(* IEC 61131-3 sources: Elmo_Master/Lasal_PRG/Welcon8Axis_EtherCAT_Test_With_RobotAxis/Network/Axis2, 1 file *)

(* ---- ONE_Axis2_Table.st ---- *)
#define OBJECTS_CONFIG

//Define part of class _LMCAxisBase
//#define _DEBUG_MODUS_MUTEX_OFF
//#define _DEBUG_MODUS_ISSYNCHRON
//#define _DEBUG_MODUS_CHECKSWLIMIT
//#define _DEBUG_MODUS_BRAKING

#define _LMCAXIS_NORMOVERRIDE         1000    // Dieser Override-Wert entspricht 100%.
#define _LMCAXIS_MAXOVERRIDE	        1000		// Maximalwert für Override im LMCAXISBASE (kann mit SetParameter verändert werden.)
#define _LMCAXIS_MINOVERRIDE	           0		// Minimalwert für Override im _LMCAxisBase --> damit man mit Minuswerten nicht in die falsche Richtung fahren kann

#define _LMCAXIS_MIN_POS       -16#07000000    // default MINPOS when INITvalue=0
#define _LMCAXIS_MAX_POS        16#07000000    // default MAXPOS when INITvalue=0

#define _LMCAXIS_OVERVFLOW_POS  16#06000000    // MAX POSITION for checking overflow

#define _LMCAXIS_INVALID_POS    16#3FFFFFFF    // Invalid position for calculating the velocity

#define _LMCAXIS_INTERVAL            10            // original = 10

#define _LMCAXIS_MAX_MASTERDELAY     7    // maximum cycles for delaying the coupling to the master

#define _LMCAXIS_RESO_CALBREMS 100

#ifndef _VOID_POS
  #define  _VOID_POS 16#7FFFFFFF
#endif

/////////////////////
// Polynom 5ten Grades
#define _LMCAXIS_Poly_Pos_A     2.5
#define _LMCAXIS_Poly_Pos_B     3.0
#define _LMCAXIS_Poly_Pos_C     1.0

#define LMC_POLYNOM_V0          0                     // CoupleGearPolynom wenn Slave steht
#define LMC_POLYNOM_V           1                     // CoupleGearPolynom wenn Slave fährt

//////////////////////
// Bewegungsrichtungen
#define _LMCAXIS_MOVE_ANY_WAY              0       // beide Richtungen
#define _LMCAXIS_MOVE_NEG_DIR              1       // nur negative Bewegungsrichtung
#define _LMCAXIS_MOVE_SHORTEST_WAY         2       // kürzester Weg (beide Richtungen)
#define _LMCAXIS_MOVE_POS_DIR              3       // nur positive Bewegungsrichtung

//////////////////////
// Mutex
#define MUTEX_NAME_MAX_LENGTH_LMCAXIS     32   //maximale Anzahl an Zeichen für den Mutexnamen
#define MUTEX_NAME_END_LENGTH_LMCAXIS      3
#define STR_MUTEX_NAME_SEPERATOR_LMCAXIS ".."

#define _LMCAXIS_WAITTIMEPOWERON           90sec    // Wartezeit bei PowerOn bis TimeOut entsteht (maximale Kommutierungszeitdauer beim DiasDrive für Linearmotoren sind 86sec)
#define _LMCAXIS_WAITTIMEPOWEROFF           1sec    // Wartezeit bei PowerOff bis TimeOut entsteht

#define _LMCAXIS_Max_V_FILTER_SIZE   100

//////////////////////
// ruckbegrenzter Modus _JERK_PROFILE
#define MIN_SHRINK_FACTOR_4_CORRECTTOEXACTPOS 0.9
#define MAX_SHRINK_FACTOR_4_CORRECTTOEXACTPOS_FAR 1.2
#define MAX_SHRINK_FACTOR_4_CORRECTTOEXACTPOS_NEAR 5.0
#define MAX_SHRINK_FACTOR_4_CORRECTTOEXACTPOS_WINDOW 5.0

#define MAX_TIME_TO_WAIT_4_BRAKING 3.0 //in Ticks
#define MAX_DURATION_WITH_MAX_ACCEL_TO_MASTER 20000  //in Ticks
#define ALLOWED_AJMP_FACTOR 1.1
#define FACTOR_4_ALLOWED_MASTER_ACCEL_PROFILE_COUPLING 1.2
#define ACCEL_FACTOR_4_PROFILE_COUPLING 1.1
#define JERK_FACTOR_4_PROFILE_COUPLING 1.2

//////////////////////
// LREAL Modi
// #define DEBUG_TRAP_DELTA_ACCEL
#define _LMCAXIS_LREAL_EPSILON 0.000001

#ifndef _DINT_MIN
#define _DINT_MIN -2147483648
#endif

#ifndef _DINT_MAX
#define _DINT_MAX 2147483647
#endif

#define _LMCAXIS_MIN_VEL_MOVECMD 1 // minimale programmierbare Geschwindigkeit fuer LREAL-MoveTypes [internal units / sec]

#define _LMCAXIS_SAFEREFERENCE_TIMEOUT          10 SEC
#define _LMCAXIS_SBTACTIVE_TIMEOUT              16 SEC
#define _LMCAXIS_SAFETYASYNCREQUEST_REPEATTIME  200 MS

#define _LMCAXIS_SBT_SAFESTATE_TESTIDLE    16#0
#define _LMCAXIS_SBT_SAFESTATE_TESTDONE    16#6
#define _LMCAXIS_SBT_SAFESTATE_ERROR      16#E0
#define _LMCAXIS_SBT_FUNCSTATE_FINISH        13

#define _LMCAXIS_LMCPROF_NEWINST_STOPMOVE    77

//+++ einbau HP 13.9.2011 +++++++++++++++++++++++++++++++++++++++++++++++++++++++

//////////////////////
// CoupleGearPolynom
#define _LMCAXIS_FACTOR_JMAX         10
#define _LMCAXIS_FACTOR_T_VAL_X      0.80
#define _LMCAXIS_FACTOR_T_VAL_Z      0.80
#define _LMCAXIS_MIN_TICKS           0

//#define REPORT_TRAPEZOIDSPLINE_DISABLED
#undef REPORT_TRAPEZOIDSPLINE_DISABLED

// Formeltest und Test auf numerische Genauigkeit
//#define CHECK_PRECISION

#define PRAEFIX_KILO          (1000.0)
#ifndef CONVERT_SEC_TO_MSEC
  #define CONVERT_SEC_TO_MSEC   (1000.0)
#endif
//+++++++++++++++++++++++++++++++++++++++++++++++++++++++ einbau HP 13.9.2011 +++

#ifndef LMCMODULEBASE_MAX_LOGININDEX
  #define LMCMODULEBASE_MAX_LOGININDEX      9
#endif

// ===================================================================
// defines linked to safety features
// defines from header file DriveSafetyIF.h from HW lib to reduce dependencies

// VERIFY CMDRSP
// General
#define _LMCAXIS_SAFETY_VERCMD_OK                     0x40000000  // Command successfully processed
#define _LMCAXIS_SAFETY_VERCMD_BUSY                   0x0000000B  // Response to command has not yet been recived
#define _LMCAXIS_SAFETY_VERCMD_EXECUTING              0x4000000B  // Commmand ist still beeing processed ins safety FW
#define _LMCAXIS_SAFETY_VERCMD_WRONG_RUNSTATE         0x40000003  // Command not allowed in current state
#define _LMCAXIS_SAFETY_VERCMD_NOT_NEEDED             0x40000004  // Command executed, although no verification is necessary

#define _LMCAXIS_SAFETY_VERCMD_ERROR_ENC_ID_PROG      0x40000005  // Programming of the encoder index failed

#define _LMCAXIS_SAFETY_VERCMD_INCOMPLETE             0x40000001  // Not all axes requiring verification, have been verified
#define _LMCAXIS_SAFETY_VERCMD_ERROR                  0x40000002  // Saving the HDSL verification status has failed

// VERIFY STATE
#define _LMCAXIS_SAFETY_VERSTATE_UNKOWN               0x00000000  // State has not yet been read
#define _LMCAXIS_SAFETY_VERSTATE_BUSY                 0x0000000B  // State is beeing read

#define _LMCAXIS_SAFETY_VERSTATE_NOT_VERIFIED         0x1A8C5E7B  // Axis not verified, verification necessary
#define _LMCAXIS_SAFETY_VERSTATE_SYSTEM_VERIFIED      0x2B9D6F8C  // Entire drive fully verified
#define _LMCAXIS_SAFETY_VERSTATE_NOT_USED             0x30000000  // no verification necessary for this axis, as not configured as Hiperface DSL

#define _LMCAXIS_SAFETY_VERSTATE_VERIFICATION_PENDING 0x30000001  // Verification has been started for this axis, Programming of the encoder index in progress
#define _LMCAXIS_SAFETY_VERSTATE_AXIS_VERIFIED        0x30000002  // Encoder index has been successfully programmed, Verification completed for this axis (Overall verification necessary at the end)

// REFERENCE CMDRSP
// General
#define _LMCAXIS_SAFETY_REFCMD_OK                     0x40000000  // Command successfully processed
#define _LMCAXIS_SAFETY_REFCMD_BUSY                   0x0000000B  // Response to command has not yet been recived
#define _LMCAXIS_SAFETY_REFCMD_PROGRAMMING_FAILED     0x40000002  // The saving of the offset or the referencing status has failed.
#define _LMCAXIS_SAFETY_REFCMD_WRONG_RUNSTATE         0x40000003  // Command not allowed in current state
#define _LMCAXIS_SAFETY_REFCMD_NOT_NEEDED             0x40000004  // Command executed, although no reference is necessary

// For _LMCAXIS_SAFETY__REFCMD_ACKZERO_POS
#define _LMCAXIS_SAFETY_REFCMD_NOT_ALLOWED            0x40000010  // Absolute position referencing was not started, command not yet allowed
#define _LMCAXIS_SAFETY_REFCMD_NO_MOVEMENT            0x40000011  // Position has not moved far enough from the zero position since the start of referencing
#define _LMCAXIS_SAFETY_REFCMD_WRONG_POSITION         0x40000012  // Newly approached zero position deviates more than permitted from initially approached zero position

// REFERENCE STATE
#define _LMCAXIS_SAFETY_REFSTATE_UNKOWN               0x00000000  //

#define _LMCAXIS_SAFETY_REFSTATE_BUSY                 0x0000000B  // State is beeing read

#define _LMCAXIS_SAFETY_STATE_NOT_REFERENCED          0x1A8C5E7B  // Axis not referenced, referencing necessary
#define _LMCAXIS_SAFETY_STATE_AXIS_REFERENCED         0x2B9D6F8C  // Axis fully referenced
#define _LMCAXIS_SAFETY_STATE_NOT_NEEDED              0x30000000  // No referencing necessary for this axis

#define _LMCAXIS_SAFETY_STATE_WAIT_MOVEMENT           0x30000001  // Referencing has been started, it is waiting for the waiting for the current position to move away from the zero position
#define _LMCAXIS_SAFETY_STATE_ACK_PENDING             0x30000002  // Current position far enough away from zero position, it waits for the zero position to be approached again and confirmed
#define _LMCAXIS_SAFETY_STATE_REFERENCE_DONE          0x30000003  // Zero position successfully confirmed, referencing completed

// DRIVE SAFETY PARA STATES
#define _LMCAXIS_SAFETY_UPDATEPARACLASS_STATE                 16#857E
#define _LMCAXIS_SAFETY_UPDATEPARACLASS_STATE_VER_1           1                   //version 1
#define _LMCAXIS_SAFETY_UPDATEPARACLASS_STATE_VER_MAX         _LMCAXIS_SAFETY_UPDATEPARACLASS_STATE_VER_1   //newest implemented version

#define _LMCAXIS_SAFETY_UPDATEPARACLASS_STATE_GENERAL_ERROR                 1
#define _LMCAXIS_SAFETY_UPDATEPARACLASS_STATE_ASYNC_BUSY                    3
#define _LMCAXIS_SAFETY_UPDATEPARACLASS_STATE_GENERAL_READY                 5
#define _LMCAXIS_SAFETY_UPDATEPARACLASS_STATE_UPDATE_CY                     6
#define _LMCAXIS_SAFETY_UPDATEPARACLASS_STATE_SAFETY_READY                  10
#define _LMCAXIS_SAFETY_UPDATEPARACLASS_STATE_SAFETY_ERROR                  11
#define _LMCAXIS_SAFETY_UPDATEPARACLASS_STATE_SAFETY_CHANGED                12
#define _LMCAXIS_SAFETY_UPDATEPARACLASS_STATE_SAFETY_SETSERVICEMODE_PENDING 20
#include <.\lsl_st_systrace.h>
#include "..\..\Class\_LMCAxisBase\C_MathAxis.h"
#include "..\..\Class\_LMCAxisBase\_LMCTraceView.h"
#include "..\..\Class\_LMCAxisBase\BacklashLogin.h"
#include "..\..\Class\_LMCAxisBase\TorqueHandlingLogin.h"
//Define part of class _LMCAxisVOVMonitoring
// Monitoring time (ms). If a button is not being pressed or released for a this amount of time the connection has been broken
#ifndef LMCAXIS_VOVMonitor_NoReactionTimeLimit
  #define  LMCAXIS_VOVMonitor_NoReactionTimeLimit 1000 ms
#endif
//Define part of class _LMCMathFunctions
#define _INT_DEG                       * 1024 * 1000 //Internal Resolution of Degrees
#define LMC_PI                          3.1415926535897932384626433832795   //LMC_ avoids name clash

#define _LMC_EPSILON    0.000001
#define _MATH_EPSILON   0.000000001

//LREAL Zero Test:
#ifndef _LMCMATH_FLOAT_ISZERO
  #define _LMCMATH_FLOAT_ISZERO(p1)            ((p1 > -_LMC_EPSILON) & (p1 < _LMC_EPSILON))
#endif
#ifndef _LMCMATH_FLOAT_NOTZERO
  #define _LMCMATH_FLOAT_NOTZERO(p1)           ((p1 < -_LMC_EPSILON) | (p1 > _LMC_EPSILON))
#endif
#ifndef _LMCMATH_FLOAT_EQUAL
  #define _LMCMATH_FLOAT_EQUAL(p1,p2)          (((p1 - p2) < _LMC_EPSILON) & ((p1 - p2) > -_LMC_EPSILON))
#endif

#define _LMCMATH_LREAL_MAX  1.79E308
#define _LMCMATH_REAL_MAX   3.4E38

#ifndef _DINT_MIN
  #define _DINT_MIN -2147483648
#endif

#define LMC_NUMERIC_TOLERANCE   (0.000000001)
#define LMC_RESOLVE_TOLERANCE       (0.000000001)

// 25µsec für ein repeat auf ARM CP 111
#define LMC_MAX_REPEAT      25

// Geschwindigkeit wird auf 1 interne Einheit genau iteriert
#define PRECIS_REPEAT   (1.0)

//#define INTERN_MATH_TEST
#include "..\..\Class\_LMCMathFunctions\C_MathFunct.h"
//Define part of class Controller
#define MaxDragDelayCycles 20

// define of NewInst index to read hardware diagnosis data from HWK
#define LMCCONTROLLER_GET_HARDWARE_DIAGNOSIS      16#83B1

// defines to mark maximum values of DINT as floating number
#ifndef LMCCONTROLLER_DINT_MIN_LREAL
  #define LMCCONTROLLER_DINT_MIN_LREAL -2147483648.0
#endif

#ifndef LMCCONTROLLER_DINT_MAX_LREAL
  #define LMCCONTROLLER_DINT_MAX_LREAL 2147483647.0
#endif

FUNCTION GLOBAL TAB ONE_Axis2
-1$UINT, 0$UINT,
0$UINT, 0$UINT,

17$UDINT,
TO_UDINT(1047453148), "_AxisBase", 1$UINT, 58$UINT, 0$UINT,
TO_UDINT(3162349954), "_LMCABSEncoder", 1$UINT, 0$UINT, 1$UINT,
TO_UDINT(1422175863), "_LMCAxis", 1$UINT, 120$UINT, 1$UINT,
TO_UDINT(280984637), "_LMCAxisBase", 2$UINT, 111$UINT, 0$UINT,
TO_UDINT(2147194214), "_LMCAxisRef", 1$UINT, 32$UINT, 1$UINT,
TO_UDINT(3113915997), "_LMCAxisVis", 1$UINT, 42$UINT, 1$UINT,
TO_UDINT(3511906983), "_LMCAxisVisInt", 1$UINT, 63$UINT, 1$UINT,
TO_UDINT(1670072687), "_LMCAxisVisLogHandle", 1$UINT, 0$UINT, 1$UINT,
TO_UDINT(4049061347), "_LMCAxisVisLogViewer", 1$UINT, 0$UINT, 5$UINT,
TO_UDINT(3953984284), "_LMCAxisVisPara", 1$UINT, 13$UINT, 1$UINT,
TO_UDINT(3513915334), "_LMCAxisVOVMonitoring", 1$UINT, 2$UINT, 1$UINT,
TO_UDINT(838927485), "_LMCMathFunctions", 1$UINT, 75$UINT, 1$UINT,
TO_UDINT(1117088251), "_LMCPublisher", 1$UINT, 0$UINT, 1$UINT,
TO_UDINT(1736530975), "_LMCRefBase", 1$UINT, 11$UINT, 0$UINT,
TO_UDINT(3213872914), "_LMCSafety", 1$UINT, 21$UINT, 1$UINT,
TO_UDINT(1198357413), "Controller", 1$UINT, 47$UINT, 0$UINT,
TO_UDINT(28504452), "PosController", 2$UINT, 77$UINT, 1$UINT,

1$UINT, TO_UDINT(1393205339), "_LMCAXIS_AXIS2\_LMCABSENCODER1",

_NO_ATTR, TO_UDINT(1250969566), "_LMCAXIS_AXIS2",

1$UINT, TO_UDINT(2274490556), "_LMCAXIS_AXIS2\_LMCAXISREF1",

1$UINT, TO_UDINT(912027803), "_LMCAXIS_AXIS2\_LMCAXISVIS1",

1$UINT, TO_UDINT(3549664169), "_LMCAXIS_AXIS2\_LMCAXISVIS1\_LMCAXISVISINT1",

1$UINT, TO_UDINT(3510254084), "_LMCAXIS_AXIS2\_LMCAXISVIS1\_LMCAXISVISLOGHANDLE1",

1$UINT, TO_UDINT(900082051), "_LMCAXIS_AXIS2\_LMCAXISVIS1\_LMCAXISVISLOGVIEWER1",
1$UINT, TO_UDINT(2897180729), "_LMCAXIS_AXIS2\_LMCAXISVIS1\_LMCAXISVISLOGVIEWER2",
1$UINT, TO_UDINT(3685238959), "_LMCAXIS_AXIS2\_LMCAXISVIS1\_LMCAXISVISLOGVIEWER3",
1$UINT, TO_UDINT(1171053836), "_LMCAXIS_AXIS2\_LMCAXISVIS1\_LMCAXISVISLOGVIEWER4",
1$UINT, TO_UDINT(852225434), "_LMCAXIS_AXIS2\_LMCAXISVIS1\_LMCAXISVISLOGVIEWER5",

1$UINT, TO_UDINT(841254793), "_LMCAXIS_AXIS2\_LMCAXISVIS1\_LMCAXISVISPARA1",

1$UINT, TO_UDINT(1593456117), "_LMCAXIS_AXIS2\_LMCAXISVIS1\_LMCAXISVOVMONITORING",

1$UINT, TO_UDINT(3529465846), "_LMCAXIS_AXIS2\_LMCMATHFUNCTIONS1",

1$UINT, TO_UDINT(2748705581), "_LMCAXIS_AXIS2\_LMCPUBLISHER1",

1$UINT, TO_UDINT(2568002256), "_LMCAXIS_AXIS2\_LMCSAFETY1",

_NO_ATTR, TO_UDINT(1207330664), "POSCONTROLLER_AXIS2",

//Internal connections
0$UDINT,
15$UDINT,
TO_UDINT(1), "_LMCMathFunctions1", TO_UDINT(13),
TO_UDINT(1), "_LMCABSEncoder1", TO_UDINT(0),
TO_UDINT(1), "_LMCAxisVis1", TO_UDINT(3),
TO_UDINT(1), "_LMCAxisRef1", TO_UDINT(2),
TO_UDINT(1), "_LMCSafety1", TO_UDINT(15),
TO_UDINT(1), "_LMCPublisher1", TO_UDINT(14),
TO_UDINT(3), "_LMCAxisVisInt1", TO_UDINT(4),
TO_UDINT(3), "_LMCAxisVisPara1", TO_UDINT(11),
TO_UDINT(3), "_LMCAxisVisLogViewer1", TO_UDINT(6),
TO_UDINT(3), "_LMCAxisVisLogViewer2", TO_UDINT(7),
TO_UDINT(3), "_LMCAxisVisLogViewer3", TO_UDINT(8),
TO_UDINT(3), "_LMCAxisVisLogViewer4", TO_UDINT(9),
TO_UDINT(3), "_LMCAxisVisLogViewer5", TO_UDINT(10),
TO_UDINT(3), "_LMCAxisVisLogHandle1", TO_UDINT(5),
TO_UDINT(3), "_LMCAxisVOVMonitoring", TO_UDINT(12),
0$UDINT,
15$UDINT,
TO_UDINT(1), "LMCController", TO_UDINT(16), "Signal_Input",
TO_UDINT(1), "LMCMath", TO_UDINT(13), "ClassSvr",
TO_UDINT(1), "LMCSafety", TO_UDINT(15), "ClassSvr",
TO_UDINT(1), "LMCReference", TO_UDINT(2), "RefInput",
TO_UDINT(1), "LMCAbsEncoder", TO_UDINT(0), "ClassSvr",
TO_UDINT(1), "LMCPublisher", TO_UDINT(14), "ClassSvr",
TO_UDINT(3), "LMCAxisBase", TO_UDINT(1), "Control",
TO_UDINT(4), "LMCAxisVisPara", TO_UDINT(11), "ClassSvr",
TO_UDINT(6), "LogIndex", TO_UDINT(5), "LogIndex",
TO_UDINT(7), "LogIndex", TO_UDINT(5), "LogIndex",
TO_UDINT(8), "LogIndex", TO_UDINT(5), "LogIndex",
TO_UDINT(9), "LogIndex", TO_UDINT(5), "LogIndex",
TO_UDINT(10), "LogIndex", TO_UDINT(5), "LogIndex",
TO_UDINT(11), "ocLMCAxisVisInt", TO_UDINT(4), "ClassSvr",
TO_UDINT(12), "ToVisInt", TO_UDINT(4), "ClassSvr",

//Initialization values
0$UDINT,
30$UDINT,
TO_UDINT(1), "SimulateMode", TO_UDINT(0),//|Axis2._LMCAxis_Axis2.SimulateMode;
TO_UDINT(1), "ExUnits", TO_UDINT(4096),//|Axis2._LMCAxis_Axis2.ExUnits;
TO_UDINT(1), "IntUnits", TO_UDINT(1 mm),//|Axis2._LMCAxis_Axis2.IntUnits;
TO_UDINT(1), "VMax", TO_UDINT(50 mm),//|Axis2._LMCAxis_Axis2.VMax;
TO_UDINT(1), "AMax", TO_UDINT(5000 mm),//|Axis2._LMCAxis_Axis2.AMax;
TO_UDINT(1), "Tjerk", TO_UDINT(0),//|Axis2._LMCAxis_Axis2.Tjerk;
TO_UDINT(1), "MoveType", TO_UDINT(_RAMP_Profile),//|Axis2._LMCAxis_Axis2.MoveType;
TO_UDINT(1), "Resolution", TO_UDINT(1),//|Axis2._LMCAxis_Axis2.Resolution;
TO_UDINT(1), "Modulo", TO_UDINT(0),//|Axis2._LMCAxis_Axis2.Modulo;
TO_UDINT(1), "SWMinPos", TO_UDINT(0),//|Axis2._LMCAxis_Axis2.SWMinPos;
TO_UDINT(1), "SWMaxPos", TO_UDINT(0),//|Axis2._LMCAxis_Axis2.SWMaxPos;
TO_UDINT(1), "ErrorConfig", TO_UDINT(2#0000000001000000),//|Axis2._LMCAxis_Axis2.ErrorConfig;
TO_UDINT(1), "AEmergency", TO_UDINT(0),//|Axis2._LMCAxis_Axis2.AEmergency;
TO_UDINT(1), "JMax", TO_UDINT(0),//|Axis2._LMCAxis_Axis2.JMax;
TO_UDINT(1), "Config", TO_UDINT(0),//|Axis2._LMCAxis_Axis2.Config;
TO_UDINT(1), "ID", TO_UDINT(0),//|Axis2._LMCAxis_Axis2.ID;
TO_UDINT(4), "TriangleMode", TO_UDINT(1),//|Axis2._LMCAxisVis1\_LMCAxis_Axis2\_LMCAxisVisInt1.TriangleMode;
TO_UDINT(6), "LogOffset", TO_UDINT(0),//|Axis2._LMCAxisVis1\_LMCAxis_Axis2\_LMCAxisVisLogViewer1.LogOffset;
TO_UDINT(7), "LogOffset", TO_UDINT(1),//|Axis2._LMCAxisVis1\_LMCAxis_Axis2\_LMCAxisVisLogViewer2.LogOffset;
TO_UDINT(8), "LogOffset", TO_UDINT(2),//|Axis2._LMCAxisVis1\_LMCAxis_Axis2\_LMCAxisVisLogViewer3.LogOffset;
TO_UDINT(9), "LogOffset", TO_UDINT(3),//|Axis2._LMCAxisVis1\_LMCAxis_Axis2\_LMCAxisVisLogViewer4.LogOffset;
TO_UDINT(10), "LogOffset", TO_UDINT(4),//|Axis2._LMCAxisVis1\_LMCAxis_Axis2\_LMCAxisVisLogViewer5.LogOffset;
TO_UDINT(11), "MovRefPosWindow", TO_UDINT(0),//|Axis2._LMCAxisVis1\_LMCAxis_Axis2\_LMCAxisVisPara1.MovRefPosWindow;
TO_UDINT(14), "Config", TO_UDINT(0),//|Axis2._LMCAxis_Axis2\_LMCPublisher1.Config;
TO_UDINT(14), "ID", TO_UDINT(0),//|Axis2._LMCAxis_Axis2\_LMCPublisher1.ID;
TO_UDINT(16), "iHWErrors", TO_UDINT(0),//|Axis2.PosController_Axis2.iHWErrors;
TO_UDINT(16), "vHWDelay", TO_UDINT(0),//|Axis2.PosController_Axis2.vHWDelay;
TO_UDINT(16), "oActive", TO_UDINT(0),//|Axis2.PosController_Axis2.oActive;
TO_UDINT(16), "cDragLimit", TO_UDINT(0),//|Axis2.PosController_Axis2.cDragLimit;
TO_UDINT(16), "cDragCalcDelay", TO_UDINT(0),//|Axis2.PosController_Axis2.cDragCalcDelay;

//Symbolic initialization values
0$UDINT,
0$UDINT,

//Initialization of string values
0$UDINT,
0$UDINT,

//Configuration of tasks (RealTime, Cyclic, Background)
0$UDINT,
1$UDINT,
TO_UDINT(1), (1)$UDINT, 4194303$DINT, 	//_LMCAXIS_AXIS2

0$UDINT,
0$UDINT,

0$UDINT,
2$UDINT,
TO_UDINT(1), (100)$UDINT, 4194303$DINT, 	//_LMCAXIS_AXIS2
TO_UDINT(12), (100)$UDINT, 4194303$DINT, 	//_LMCAXIS_AXIS2\_LMCAXISVIS1\_LMCAXISVOVMONITORING

//External connections
0$UDINT,
8$UDINT,
TO_UDINT(1), "ActPosition", C_TRY, TO_UDINT(4273818432), "DriveAxisDS402_Axis2","ActPos",
TO_UDINT(1), "HWReady", C_TRY, TO_UDINT(3391823300), "WELCON_11","Online",
TO_UDINT(1), "HWError", C_TRY, TO_UDINT(4273818432), "DriveAxisDS402_Axis2","AxError",
TO_UDINT(16), "iHWErrors", C_TRY, TO_UDINT(4273818432), "DriveAxisDS402_Axis2","AxError",
TO_UDINT(16), "oActive", C_TRY, TO_UDINT(4273818432), "DriveAxisDS402_Axis2","AxEnable",
TO_UDINT(16), "oOutputSignal", C_TRY, TO_UDINT(4273818432), "DriveAxisDS402_Axis2","SetPos",
TO_UDINT(16), "DriveEnabled", C_TRY, TO_UDINT(4273818432), "DriveAxisDS402_Axis2","AxEnable",
TO_UDINT(16), "HWErrorQuit", C_TRY, TO_UDINT(4273818432), "DriveAxisDS402_Axis2","AxErrorQuit",

//Magic internal connections
0$UDINT,
21$UDINT,
TO_UDINT(2), "HWMin", TO_UDINT(1), "HWMin",
TO_UDINT(2), "HWMax", TO_UDINT(1), "HWMax",
TO_UDINT(2), "ZImpulse", TO_UDINT(1), "ZImpulse",
TO_UDINT(2), "RefSwitch", TO_UDINT(1), "RefSwitch",
TO_UDINT(2), "LatchPos", TO_UDINT(1), "LatchPos",
TO_UDINT(4), "LMCAxisBase", TO_UDINT(3), "LMCAxisBase",
TO_UDINT(5), "LMCAxisBase", TO_UDINT(3), "LMCAxisBase",
TO_UDINT(6), "LMCAxisBase", TO_UDINT(3), "LMCAxisBase",
TO_UDINT(7), "LMCAxisBase", TO_UDINT(3), "LMCAxisBase",
TO_UDINT(8), "LMCAxisBase", TO_UDINT(3), "LMCAxisBase",
TO_UDINT(9), "LMCAxisBase", TO_UDINT(3), "LMCAxisBase",
TO_UDINT(10), "LMCAxisBase", TO_UDINT(3), "LMCAxisBase",
TO_UDINT(14), "Provider", TO_UDINT(1), "Provider",
TO_UDINT(14), "Config", TO_UDINT(1), "Config",
TO_UDINT(14), "ID", TO_UDINT(1), "ID",
TO_UDINT(15), "HWReady", TO_UDINT(1), "HWReady",
TO_UDINT(15), "HWError", TO_UDINT(1), "HWError",
TO_UDINT(15), "HWMin", TO_UDINT(1), "HWMin",
TO_UDINT(15), "HWMax", TO_UDINT(1), "HWMax",
TO_UDINT(15), "Emergency", TO_UDINT(1), "Emergency",
TO_UDINT(15), "LMCController", TO_UDINT(1), "LMCController",

//Configuration of timeslots of tasks (RealTime, Cyclic)
#ifdef __LSLLDR_TIMESLOTS__
0$UDINT,
0$UDINT,

0$UDINT,
0$UDINT,

#endif //__LSLLDR_TIMESLOTS__

//MultiMaster connections
#ifdef __LSLLDR_MULTIMASTER__
0$UDINT,
0$UDINT,
#endif //__LSLLDR_MULTIMASTER__

//Configuration for task ID (RealTime, CyclicTime)
#ifdef __LSLLDR_TASKID__
"\\\\TASKS2  "
0$UDINT,
1$UDINT,
(0)$UDINT, 	//_LMCAXIS_AXIS2

0$UDINT,
0$UDINT,

0$UDINT,
2$UDINT,
(0)$UDINT, 	//_LMCAXIS_AXIS2
(0)$UDINT, 	//_LMCAXIS_AXIS2\_LMCAXISVIS1\_LMCAXISVOVMONITORING

#endif //__LSLLDR_TASKID__

END_FUNCTION
